Fanuc KAREL source: KT00598.KL

PROGRAM KT00598
%NOLOCKGROUP
VAR
  I1: INTEGER
  I2: INTEGER
  OUT: INTEGER
BEGIN
  I1 = 2
  I2 = 3
  I1 = 2
  I2 = 3
  OUT = NOT I1
END KT00598
